(* IEC 61131-3 sources: sis-interlock-demo/tests/POUs/Helpers/FB_SisHarness, 6 files *)

(* ---- FB_SisHarness.decl.st ---- *)
// Назначение: стенд сценарных тестов по матрице (DESIGN.md, 12.5): настоящие FB_SisApp, GVL_SisCfg
//             и ST_SisIo с подменным временем PL.FB_FakeTime и журналом FB_SisEventLog — от тегов на
//             входе до тегов на выходе, как на FAT. Тесты пишут stIo и stCmd по имени экземпляра
//             (они во VAR_INPUT: запись в VAR извне — ошибка C0037) и читают fbApp, fbLog.
// Автор:      kr0nsch
// Версия:     0.1.0
// Документ:   docs/DESIGN.md, раздел «12.5 Стенд FB_SisHarness»
// ВНИМАНИЕ:   код демонстрационный и не предназначен для систем безопасности. Реальная ПАЗ
//             требует определения SIL, сертифицированных аппаратных и программных средств
//             и валидации по ГОСТ Р МЭК 61511.
FUNCTION_BLOCK FB_SisHarness
VAR_INPUT
    stIo  : ST_SisIo;              // образ ввода-вывода: тест ставит входы, читает выходы xQ*
    stCmd : ST_SisCmd;             // команды HMI: сброс, пусковые обходы, байпасы
END_VAR
VAR
    fbTime  : PL.FB_FakeTime;      // подменное время, старт LTIME#1H
    fbLog   : FB_SisEventLog;      // журнал событий ПАЗ
    fbApp   : FB_SisApp;           // ПАЗ объекта под тестом
    udiMark : UDINT;               // номер последнего события на момент MarkEvents
END_VAR
VAR CONSTANT
    RUN_MAX_ITERATIONS : UINT := 1500;   // предел шагов одного Run: все тесты идут в одном цикле задачи
END_VAR

(* ---- HasEvent.method.decl.st ---- *)
// TRUE — после MarkEvents в журнале есть событие eKind причины uiCause (порядок внутри вызова не важен).
METHOD HasEvent : BOOL
VAR_INPUT
    eKind   : E_SisEventKind;   // вид события
    uiCause : UINT;             // номер причины
END_VAR
VAR
    uiBack : UINT;              // сколько событий назад
    stEv   : ST_SisEvent;       // событие журнала
    xNewer : BOOL;              // событие новее отметки
END_VAR

(* ---- Keys.method.decl.st ---- *)
// Ключи разрешения байпасов и пусковых обходов; кнопка «Сброс ПАЗ» отпущена. Цикл не выполняется.
METHOD Keys
VAR_INPUT
    xBypass   : BOOL;   // ключ «Разрешение байпасов»
    xOverride : BOOL;   // ключ «Разрешение пусковых обходов»
END_VAR

(* ---- Run.method.decl.st ---- *)
// Шаги tStep до суммарной длительности tDuration, последний шаг — остаток; tDuration = T#0S — ничего;
// tStep = T#0S — один шаг на всю длительность. Не больше RUN_MAX_ITERATIONS шагов.
METHOD Run
VAR_INPUT
    tDuration : TIME;   // сколько времени прогнать
    tStep     : TIME;   // шаг
END_VAR
VAR
    tLeft  : TIME;      // осталось
    tThis  : TIME;      // шаг этой итерации
    uiIter : UINT;      // итераций
END_VAR

(* ---- Run.method.impl.st ---- *)
tLeft := tDuration;
uiIter := 0;
WHILE tLeft > T#0S AND uiIter < RUN_MAX_ITERATIONS DO
    IF tStep > T#0S AND tStep < tLeft THEN
        tThis := tStep;
    ELSE
        tThis := tLeft;
    END_IF
    Step(tStep := tThis);
    tLeft := tLeft - tThis;
    uiIter := uiIter + 1;
END_WHILE

(* ---- Step.method.decl.st ---- *)
// Шаг времени и цикл ПАЗ.
METHOD Step
VAR_INPUT
    tStep : TIME;   // шаг подменного времени
END_VAR
